// TIA Portal V20 export
// export: Created 2026-10-11T05:32:37.9298943Z, ExportSetting WithDefaults, DisplayName Totally Integrated Automation Portal, DisplayVersion V20, DisplayName TIA Portal Openness, DisplayVersion V20, DisplayName TIA Portal Teamcenter Gateway, DisplayVersion V20, DisplayName TIA Portal Version Control Interface, DisplayVersion V20, DisplayName SINAMICS Startdrive Advanced, DisplayVersion V20 SP1 Update 2, DisplayName SINAMICS Startdrive G110M, G120, G120C, G120D, G120P, G115D, DisplayVersion V20 SP1 Update 2, DisplayName SINAMICS Startdrive G130, G150, S120, S150, SINAMICS MV, G220, S200, S210, DisplayVersion V20 SP1 Update 2, DisplayName STEP 7 Professional, DisplayVersion V20, DisplayName STEP 7 Safety, DisplayVersion V20, DisplayName WinCC Basic/Comfort/Advanced, DisplayVersion V20, DisplayName WinCC Professional, DisplayVersion V20, DisplayName WinCC Unified, DisplayVersion V20
FUNCTION "FRK_UnitFinish" : Void   // FC51, SCL
{ S7_Optimized_Access := 'TRUE' }
VERSION : 0.1
// stored: AutoNumber true, IsIECCheckEnabled false, SetENOAutomatically false, UDAEnableTagReadback false
   VAR_IN_OUT
      Core : "FRK_Core";
      Unit : "FRK_Unit";
      Response : "ST_HmiResponse";
      Status : "ST_ModuleStatus";
      Part : "ST_PartContext";
      History : Array[1..16] of "ST_Diagnostic";
      Head : Int;
   END_VAR
BEGIN

   IF #Core.Exec = 3 THEN
       IF NOT #Unit.EvReset THEN
           #Unit.FaultLatched := TRUE;
       END_IF;
       IF NOT #Unit.PrevError THEN
           "FRK_PartAborted"(Core := #Core,
                             Unit := #Unit,
                             Status := #Status,
                             Part := #Part,
                             History := #History,
                             Head := #Head);
       END_IF;
   END_IF;
   #Unit.PrevError := #Core.Exec = 3;
   IF #Core.Exec = 2 OR #Core.Exec = 4 THEN
       #Unit.RunReq := FALSE;
   END_IF;
   IF #Unit.Clearing AND #Core.Exec = 0 THEN
       IF "FRK_DescendantsReady"(OwnerIndex := #Core.RegIndex) THEN
           #Unit.Clearing := FALSE;
       END_IF;
   END_IF;
   #Unit.AbortReq := FALSE;
   #Unit.ReleaseChildren := FALSE;
   #Unit.EvReset := FALSE;
   IF #Unit.RequestPending THEN
       #Response.AckSequence := #Unit.SeenSequence;
       #Unit.RequestPending := FALSE;
   END_IF;
END_FUNCTION
